Fanuc KAREL source: KO00019.KL

PROGRAM KO00019
%NOLOCKGROUP
VAR
  P1: XYZWPREXT
  P2: XYZWPREXT
  P3: XYZWPREXT
  OUT: XYZWPREXT
BEGIN
  OUT = FRAME(P1, P2, P3)
END KO00019
